ABB RAPID module: MAIN_1.mod

MODULE MAIN_1
GLOBAL VAR robtarget robpoint0 = p:{{1015.000, 0.000, 1372.000}, {0.707107, 0.000000, 0.707107, 0.000000}, 0}{cfg 0, 0, -1, 0, 0, -1, 0, 0}{Ej 0,0,0,0,0,0}
GLOBAL VAR robtarget robpoint1 = p:{{1015.000, 0.000, 1272.000}, {0.707107, 0.000000, 0.707107, 0.000000}, 0}{cfg 0, 0, -1, 0, -1, 0, 0, 1}{Ej 0,0,0,0,0,0}
GLOBAL VAR robtarget robpoint2 = p:{{187.264, 125.487, 305.356}, {0.001606, 0.000000, 0.999999, -0.000000}, 0}{cfg -1, 0, -1, 0, 0, -1, 0, 0}{Ej 0,0,0,0,0,0}
GLOBAL VAR robtarget robpoint3 = p:{{187.786, 125.499, 139.112}, {0.001571, -0.000026, 0.999999, 0.000035}, 0}{cfg -1, 0, -1, 0, 0, -1, 0, 0}{Ej 0,0,0,0,0,0}
GLOBAL VAR robtarget robpoint4 = p:{{187.272, 447.522, 305.347}, {0.001614, 0.000009, 0.999999, -0.000017}, 0}{cfg -1, 0, 0, 0, 0, -1, 0, 0}{Ej 0,0,0,0,0,0}
GLOBAL VAR robtarget robpoint5 = p:{{187.851, 447.517, 126.235}, {0.001614, 0.000009, 0.999999, -0.000017}, 0}{cfg -1, 0, 0, 0, 0, -1, 0, 0}{Ej 0,0,0,0,0,0}
GLOBAL VAR robtarget robpoint6 = p:{{187.272, 447.522, 305.347}, {0.001614, 0.000009, 0.999999, -0.000017}, 0}{cfg -1, 0, 0, 0, 0, -1, 0, 0}{Ej 0,0,0,0,0,0}
GLOBAL VAR robtarget robpoint7 = p:{{312.208, 292.214, 255.156}, {0.086206, -0.385314, 0.917581, 0.046341}, 0}{cfg 0, 0, 0, 0, 0, -2, 0, 0}{Ej 0,0,0,0,0,0}
GLOBAL VAR robtarget robpoint8 = p:{{430.047, 43.774, 231.503}, {0.086206, -0.385314, 0.917581, 0.046341}, 0}{cfg 0, 0, -1, 0, 0, -2, 0, 0}{Ej 0,0,0,0,0,0}
GLOBAL VAR robtarget robpoint9 = p:{{109.688, -153.222, 161.073}, {0.086206, -0.385314, 0.917581, 0.046341}, 0}{cfg 0, 0, 0, 0, 0, -2, 0, 0}{Ej 0,0,0,0,0,0}
GLOBAL VAR robtarget robpoint10 = p:{{312.208, 292.214, 255.156}, {0.086206, -0.385314, 0.917581, 0.046341}, 0}{cfg 0, 0, 0, 0, 0, -2, 0, 0}{Ej 0,0,0,0,0,0}
GLOBAL VAR robtarget robpoint11 = p:{{19.898, 201.357, 302.721}, {0.032125, 0.675431, -0.735891, 0.034999}, 0}{cfg 0, 0, -1, -1, 0, 0, 0, 0}{Ej 0,0,0,0,0,0}
GLOBAL VAR robtarget robpoint12 = p:{{19.898, 174.307, 19.008}, {0.032125, 0.675431, -0.735891, 0.034999}, 0}{cfg 0, 0, 0, -1, 0, 0, 0, 0}{Ej 0,0,0,0,0,0}
GLOBAL VAR robtarget robpoint13 = p:{{378.402, 174.416, 18.997}, {0.032125, 0.675431, -0.735891, 0.034999}, 0}{cfg 0, 0, -1, 0, 0, -1, 0, 0}{Ej 0,0,0,0,0,0}
GLOBAL VAR robtarget robpoint14 = p:{{380.996, 112.363, 34.882}, {0.106872, 0.666888, -0.728163, 0.116691}, 0}{cfg 0, 0, 0, -1, 0, -1, 0, 0}{Ej 0,0,0,0,0,0}
GLOBAL VAR robtarget robpoint15 = p:{{16.551, 114.359, 34.226}, {0.106872, 0.666888, -0.728163, 0.116691}, 0}{cfg 0, 0, 0, -1, 0, 0, 0, 0}{Ej 0,0,0,0,0,0}
GLOBAL VAR robtarget robpoint16 = p:{{26.434, 54.524, 46.072}, {0.025638, -0.672233, 0.739358, 0.028195}, 0}{cfg 0, 0, 0, -1, 0, 0, 0, 0}{Ej 0,0,0,0,0,0}
GLOBAL VAR robtarget robpoint17 = p:{{385.448, 48.050, 45.137}, {0.065816, -0.669242, 0.736571, 0.072433}, 0}{cfg 0, 0, 0, 0, 0, -1, 0, 0}{Ej 0,0,0,0,0,0}
GLOBAL VAR robtarget robpoint18 = p:{{385.448, -1.625, 295.251}, {0.065816, -0.669242, 0.736571, 0.072433}, 0}{cfg 0, 0, 0, 0, 0, -1, 0, 0}{Ej 0,0,0,0,0,0}
GLOBAL VAR robtarget robpoint19 = p:{{-49.939, 252.644, 419.997}, {0.002333, -0.707103, 0.707104, 0.002024}, 0}{cfg -1, 0, 0, 0, 0, -2, 0, 0}{Ej 0,0,0,0,0,0}
GLOBAL VAR robtarget robpoint20 = p:{{-49.895, 253.259, 319.999}, {0.002333, -0.707103, 0.707104, 0.002024}, 0}{cfg -1, 0, 0, 0, 0, -2, 0, 0}{Ej 0,0,0,0,0,0}
GLOBAL VAR robtarget robpoint21 = p:{{0.000, 250.000, 270.000}, {0.002333, -0.707103, 0.707104, 0.002024}, 0}{cfg -1, 0, 0, 0, 0, -2, 0, 0}{Ej 0,0,0,0,0,0}
GLOBAL VAR robtarget robpoint22 = p:{{35.579, 247.455, 270.000}, {0.002592, -0.707102, 0.707105, 0.001666}, 0}{cfg -1, 0, 0, 0, 0, -2, 0, 0}{Ej 0,0,0,0,0,0}
GLOBAL VAR robtarget robpoint23 = p:{{70.433, 239.873, 270.000}, {0.002808, -0.707107, 0.707099, 0.001277}, 0}{cfg -1, 0, 0, 0, 0, -2, 0, 0}{Ej 0,0,0,0,0,0}
GLOBAL VAR robtarget robpoint24 = p:{{103.854, 227.408, 270.000}, {0.002956, -0.707107, 0.707100, 0.000870}, 0}{cfg -1, 0, 0, 0, 0, -2, 0, 0}{Ej 0,0,0,0,0,0}
GLOBAL VAR robtarget robpoint25 = p:{{135.160, 210.313, 270.000}, {0.003054, -0.707106, 0.707100, 0.000438}, 0}{cfg -1, 0, 0, 0, 0, -2, 0, 0}{Ej 0,0,0,0,0,0}
GLOBAL VAR robtarget robpoint26 = p:{{163.715, 188.937, 270.000}, {0.003085, -0.707106, 0.707101, 0.000000}, 0}{cfg -1, 0, 0, 0, 0, -2, 0, 0}{Ej 0,0,0,0,0,0}
GLOBAL VAR robtarget robpoint27 = p:{{188.937, 163.715, 270.000}, {0.003054, -0.707106, 0.707100, -0.000438}, 0}{cfg -1, 0, 0, 0, 0, -2, 0, 0}{Ej 0,0,0,0,0,0}
GLOBAL VAR robtarget robpoint28 = p:{{210.313, 135.160, 270.000}, {0.002968, -0.707107, 0.707100, -0.000870}, 0}{cfg -1, 0, 0, 0, 0, -2, 0, 0}{Ej 0,0,0,0,0,0}
GLOBAL VAR robtarget robpoint29 = p:{{227.408, 103.854, 270.000}, {0.002814, -0.707107, 0.707099, -0.001284}, 0}{cfg -1, 0, 0, 0, 0, -2, 0, 0}{Ej 0,0,0,0,0,0}
GLOBAL VAR robtarget robpoint30 = p:{{239.873, 70.433, 270.000}, {0.002598, -0.707102, 0.707105, -0.001672}, 0}{cfg -1, 0, 0, 0, 0, -2, 0, 0}{Ej 0,0,0,0,0,0}
GLOBAL VAR robtarget robpoint31 = p:{{247.455, 35.579, 270.000}, {0.002333, -0.707103, 0.707104, -0.002024}, 0}{cfg -1, 0, 0, 0, 0, -2, 0, 0}{Ej 0,0,0,0,0,0}
GLOBAL VAR robtarget robpoint32 = p:{{250.000, 0.000, 270.000}, {0.002024, -0.707104, 0.707103, -0.002333}, 0}{cfg -1, 0, 0, 0, 0, -2, 0, 0}{Ej 0,0,0,0,0,0}
GLOBAL VAR robtarget robpoint33 = p:{{247.455, -35.579, 270.000}, {0.001672, -0.707105, 0.707102, -0.002598}, 0}{cfg -1, 0, 0, 0, 0, -2, 0, 0}{Ej 0,0,0,0,0,0}
GLOBAL VAR robtarget robpoint34 = p:{{239.873, -70.433, 270.000}, {0.001284, -0.707099, 0.707107, -0.002814}, 0}{cfg -2, 0, 0, 0, 0, -2, 0, 0}{Ej 0,0,0,0,0,0}
GLOBAL VAR robtarget robpoint35 = p:{{227.408, -103.854, 270.000}, {0.000870, -0.707100, 0.707107, -0.002968}, 0}{cfg -2, 0, 0, 0, 0, -2, 0, 0}{Ej 0,0,0,0,0,0}
GLOBAL VAR robtarget robpoint36 = p:{{210.313, -135.160, 270.000}, {0.000438, -0.707100, 0.707106, -0.003054}, 0}{cfg -2, 0, 0, 0, 0, -2, 0, 0}{Ej 0,0,0,0,0,0}
GLOBAL VAR robtarget robpoint37 = p:{{188.937, -163.715, 270.000}, {0.000000, -0.707101, 0.707106, -0.003085}, 0}{cfg -2, 0, 0, 0, 0, -2, 0, 0}{Ej 0,0,0,0,0,0}
GLOBAL VAR robtarget robpoint38 = p:{{163.715, -188.937, 270.000}, {0.000438, 0.707100, -0.707106, 0.003054}, 0}{cfg -2, 0, 0, 0, 0, -2, 0, 0}{Ej 0,0,0,0,0,0}
GLOBAL VAR robtarget robpoint39 = p:{{135.160, -210.313, 270.000}, {0.000870, 0.707100, -0.707107, 0.002968}, 0}{cfg -2, 0, 0, 0, 0, -2, 0, 0}{Ej 0,0,0,0,0,0}
GLOBAL VAR robtarget robpoint40 = p:{{103.854, -227.408, 270.000}, {0.001284, 0.707099, -0.707107, 0.002814}, 0}{cfg -2, 0, 0, 0, 0, -2, 0, 0}{Ej 0,0,0,0,0,0}
GLOBAL VAR robtarget robpoint41 = p:{{70.433, -239.873, 270.000}, {0.001672, 0.707105, -0.707102, 0.002598}, 0}{cfg -2, 0, 0, 0, 0, -2, 0, 0}{Ej 0,0,0,0,0,0}
GLOBAL VAR robtarget robpoint42 = p:{{35.579, -247.455, 270.000}, {0.002024, 0.707104, -0.707103, 0.002333}, 0}{cfg -2, 0, 0, 0, 0, -2, 0, 0}{Ej 0,0,0,0,0,0}
GLOBAL VAR robtarget robpoint43 = p:{{0.000, -250.000, 270.000}, {0.002024, 0.707104, -0.707103, 0.002333}, 0}{cfg -2, 0, 0, 0, 0, -2, 0, 0}{Ej 0,0,0,0,0,0}
GLOBAL VAR robtarget robpoint44 = p:{{0.000, -250.000, 270.000}, {0.002333, 0.707103, -0.707104, 0.002024}, 0}{cfg -2, 0, 0, 0, 0, -2, 0, 0}{Ej 0,0,0,0,0,0}
GLOBAL VAR robtarget robpoint45 = p:{{-35.579, -247.455, 270.000}, {0.002598, 0.707102, -0.707105, 0.001672}, 0}{cfg -2, 0, 0, 0, 0, -2, 0, 0}{Ej 0,0,0,0,0,0}
GLOBAL VAR robtarget robpoint46 = p:{{-70.433, -239.873, 270.000}, {0.002808, 0.707107, -0.707099, 0.001277}, 0}{cfg -2, 0, 0, 0, 0, -2, 0, 0}{Ej 0,0,0,0,0,0}
GLOBAL VAR robtarget robpoint47 = p:{{-103.854, -227.408, 270.000}, {0.002956, 0.707107, -0.707100, 0.000870}, 0}{cfg -2, 0, 0, 0, 0, -2, 0, 0}{Ej 0,0,0,0,0,0}
GLOBAL VAR robtarget robpoint48 = p:{{-135.160, -210.313, 270.000}, {0.003054, 0.707106, -0.707100, 0.000438}, 0}{cfg -2, 0, 0, 0, 0, -2, 0, 0}{Ej 0,0,0,0,0,0}
GLOBAL VAR robtarget robpoint49 = p:{{-163.715, -188.937, 270.000}, {0.003085, 0.707106, -0.707101, 0.000000}, 0}{cfg -2, 0, 0, 0, 0, -2, 0, 0}{Ej 0,0,0,0,0,0}
GLOBAL VAR robtarget robpoint50 = p:{{-188.937, -163.715, 270.000}, {0.003054, 0.707106, -0.707100, -0.000438}, 0}{cfg -2, 0, 0, 0, 0, -2, 0, 0}{Ej 0,0,0,0,0,0}
GLOBAL VAR robtarget robpoint51 = p:{{-210.313, -135.160, 270.000}, {0.002956, 0.707107, -0.707100, -0.000870}, 0}{cfg -2, 0, 0, 0, 0, -2, 0, 0}{Ej 0,0,0,0,0,0}
GLOBAL VAR robtarget robpoint52 = p:{{-227.408, -103.854, 270.000}, {0.002801, 0.707107, -0.707099, -0.001284}, 0}{cfg -2, 0, 0, 0, 0, -2, 0, 0}{Ej 0,0,0,0,0,0}
GLOBAL VAR robtarget robpoint53 = p:{{-239.873, -70.433, 270.000}, {0.002598, 0.707102, -0.707105, -0.001672}, 0}{cfg -2, 0, 0, 0, 0, -2, 0, 0}{Ej 0,0,0,0,0,0}
GLOBAL VAR robtarget robpoint54 = p:{{-247.455, -35.579, 270.000}, {0.002333, 0.707103, -0.707104, -0.002024}, 0}{cfg -1, 0, 0, 0, 0, -2, 0, 0}{Ej 0,0,0,0,0,0}
GLOBAL VAR robtarget robpoint55 = p:{{-250.000, 0.000, 270.000}, {0.002024, 0.707104, -0.707103, -0.002333}, 0}{cfg -1, 0, 0, 0, 0, -2, 0, 0}{Ej 0,0,0,0,0,0}
GLOBAL VAR robtarget robpoint56 = p:{{-247.455, 35.579, 270.000}, {0.001666, 0.707105, -0.707102, -0.002592}, 0}{cfg -1, 0, 0, 0, 0, -2, 0, 0}{Ej 0,0,0,0,0,0}
GLOBAL VAR robtarget robpoint57 = p:{{-239.873, 70.433, 270.000}, {0.001284, 0.707099, -0.707107, -0.002801}, 0}{cfg -1, 0, 0, 0, 0, -2, 0, 0}{Ej 0,0,0,0,0,0}
GLOBAL VAR robtarget robpoint58 = p:{{-227.408, 103.854, 270.000}, {0.000870, 0.707100, -0.707107, -0.002968}, 0}{cfg -1, 0, 0, 0, 0, -2, 0, 0}{Ej 0,0,0,0,0,0}
GLOBAL VAR robtarget robpoint59 = p:{{-210.313, 135.160, 270.000}, {0.000438, 0.707100, -0.707106, -0.003054}, 0}{cfg -1, 0, 0, 0, 0, -2, 0, 0}{Ej 0,0,0,0,0,0}
GLOBAL VAR robtarget robpoint60 = p:{{-188.937, 163.715, 270.000}, {0.000000, -0.707101, 0.707106, 0.003085}, 0}{cfg -1, 0, 0, 0, 0, -2, 0, 0}{Ej 0,0,0,0,0,0}
GLOBAL VAR robtarget robpoint61 = p:{{-163.715, 188.937, 270.000}, {0.000438, -0.707100, 0.707106, 0.003054}, 0}{cfg -1, 0, 0, 0, 0, -2, 0, 0}{Ej 0,0,0,0,0,0}
GLOBAL VAR robtarget robpoint62 = p:{{-135.160, 210.313, 270.000}, {0.000870, -0.707100, 0.707107, 0.002956}, 0}{cfg -1, 0, 0, 0, 0, -2, 0, 0}{Ej 0,0,0,0,0,0}
GLOBAL VAR robtarget robpoint63 = p:{{-103.854, 227.408, 270.000}, {0.001284, -0.707099, 0.707107, 0.002814}, 0}{cfg -1, 0, 0, 0, 0, -2, 0, 0}{Ej 0,0,0,0,0,0}
GLOBAL VAR robtarget robpoint64 = p:{{-70.433, 239.873, 270.000}, {0.001672, -0.707105, 0.707102, 0.002598}, 0}{cfg -1, 0, 0, 0, 0, -2, 0, 0}{Ej 0,0,0,0,0,0}
GLOBAL VAR robtarget robpoint65 = p:{{-35.579, 247.455, 270.000}, {0.002024, -0.707104, 0.707103, 0.002333}, 0}{cfg -1, 0, 0, 0, 0, -2, 0, 0}{Ej 0,0,0,0,0,0}
GLOBAL VAR robtarget robpoint66 = p:{{0.000, 250.000, 270.000}, {0.002024, -0.707104, 0.707103, 0.002333}, 0}{cfg -1, 0, 0, 0, 0, -2, 0, 0}{Ej 0,0,0,0,0,0}
GLOBAL VAR robtarget robpoint67 = p:{{49.895, 253.258, 319.999}, {0.002024, -0.707104, 0.707103, 0.002333}, 0}{cfg -1, 0, 0, 0, 0, -2, 0, 0}{Ej 0,0,0,0,0,0}
GLOBAL VAR robtarget robpoint68 = p:{{49.939, 252.642, 419.997}, {0.002024, -0.707104, 0.707103, 0.002333}, 0}{cfg -1, 0, 0, 0, 0, -2, 0, 0}{Ej 0,0,0,0,0,0}
GLOBAL VAR robtarget robpoint69 = p:{{187.264, 125.487, 305.356}, {0.001606, 0.000000, 0.999999, -0.000000}, 0}{cfg -1, 0, -1, 0, 0, -1, 0, 0}{Ej 0,0,0,0,0,0}
GLOBAL VAR robtarget robpoint70 = p:{{187.786, 125.499, 139.112}, {0.001571, -0.000026, 0.999999, 0.000035}, 0}{cfg -1, 0, -1, 0, 0, -1, 0, 0}{Ej 0,0,0,0,0,0}
GLOBAL VAR robtarget robpoint71 = p:{{187.264, 125.487, 305.356}, {0.001606, 0.000000, 0.999999, -0.000000}, 0}{cfg -1, 0, -1, 0, 0, -1, 0, 0}{Ej 0,0,0,0,0,0}

GLOBAL VAR robtarget robpoint72 = p:{{1015.000, -1000.000, 1237.000}, {0.707107, 0.000000, 0.707107, -0.000000}, 0}{cfg -1, 0, 0, 0, 0, -1, 0, 0}{Ej 0,0,0,0,0,0}

GLOBAL Proc main()
    MoveJ robpoint0,v50,z50,tool03,wobj16
    MoveL robpoint1,v50,z50,tool03,wobj16
    SetDO D_OUT_5, 1;
    SetDO D_OUT_5, 1;
    SetDO D_OUT_5, 0.5;
    SetDO D_OUT_5, true;
    SetDO D_OUT_5, 1;
    SetDO D_OUT_5, 1;
    SetDO D_OUT_5, 0.5;
    SetDO D_OUT_5, true;
    SetDO var, val;
    SetDO var, val;
    WaitDI D_IN_5, 1;
    WaitDI D_IN_5, 1;
    WaitDI D_IN_5, 0.5;
    WaitDI D_IN_5, true;
    WaitDI D_IN_5, 1, \MaxTime:=0.1;
    WaitDI var, val;
    WaitDI var, val, \MaxTime:=0.1;
    TPWrite "Message";
    REMOTE_PROG_CALL_171;
    CODE_INSERT_172
    wobj16.x = 719.013
    wobj16.y = -664.003
    wobj16.z = 0.000
    wobj16.q1 = 1.000000
    wobj16.q2 = 0.000000
    wobj16.q3 = 0.000000
    wobj16.q4 = 0.000000
    tool03.x = 129.073
    tool03.y = 0.000
    tool03.z = 85.477
    tool03.q1 = 0.980187
    tool03.q2 = 0.000000
    tool03.q3 = 0.198076
    tool03.q4 = 0.000000
    MoveJ robpoint2,v50,z10,tool03,wobj16
    MoveL robpoint3,v100,fine,tool03,wobj16
    SetDO D_OUT_5, 1;
    PICK_PART_111;
    MoveL robpoint4,v300,z10,tool03,wobj16
    MoveL robpoint5,v100,fine,tool03,wobj16
    SetDO D_OUT_5, 0;
    PLACE_PART_112;
    MoveL robpoint6,v100,z10,tool03,wobj16
    wobj16.x = 577.67
    wobj16.y = 392.250
    wobj16.z = 0.000
    wobj16.q1 = 0.942759
    wobj16.q2 = 0.000000
    wobj16.q3 = 0.000000
    wobj16.q4 = 0.333474
    MoveJ robpoint7,v100,z25,tool03,wobj16
    MoveC robpoint8,robpoint9,v100,z25,tool03,wobj16
    MoveL robpoint10,v100,fine,tool03,wobj16
    wobj16.x = 0
    wobj16.y = 782.714
    wobj16.z = 377.610
    wobj16.q1 = 1.000000
    wobj16.q2 = 0.000000
    wobj16.q3 = 0.000000
    wobj16.q4 = 0.000000
    MoveJ robpoint11,v100,fine,tool03,wobj16
    MoveL robpoint12,v100,fine,tool03,wobj16
    MoveL robpoint13,v100,fine,tool03,wobj16
    MoveL robpoint14,v100,fine,tool03,wobj16
    MoveL robpoint15,v100,fine,tool03,wobj16
    MoveL robpoint16,v100,fine,tool03,wobj16
    MoveL robpoint17,v100,fine,tool03,wobj16
    MoveL robpoint18,v100,fine,tool03,wobj16
    EVENT_PROG_START_101;
    wobj16.x = 13.637
    wobj16.y = -840.080
    wobj16.z = 0.000
    wobj16.q1 = 0.707107
    wobj16.q2 = 0.000000
    wobj16.q3 = 0.000000
    wobj16.q4 = -0.707107
    MoveJ robpoint19,v1000,z1,tool03,wobj16
    EVENT_PATH_APPROACH_102;
    MoveL robpoint20,v1000,z1,tool03,wobj16
    MoveL robpoint21,v1000,z1,tool03,wobj16
    EVENT_PATH_START_103;
    MoveL robpoint22,v50,z1,tool03,wobj16
    MoveL robpoint23,v50,z1,tool03,wobj16
    MoveL robpoint24,v50,z1,tool03,wobj16
    MoveL robpoint25,v50,z1,tool03,wobj16
    MoveL robpoint26,v50,z1,tool03,wobj16
    MoveL robpoint27,v50,z1,tool03,wobj16
    MoveL robpoint28,v50,z1,tool03,wobj16
    MoveL robpoint29,v50,z1,tool03,wobj16
    MoveL robpoint30,v50,z1,tool03,wobj16
    MoveL robpoint31,v50,z1,tool03,wobj16
    MoveL robpoint32,v50,z1,tool03,wobj16
    MoveL robpoint33,v50,z1,tool03,wobj16
    MoveL robpoint34,v50,z1,tool03,wobj16
    MoveL robpoint35,v50,z1,tool03,wobj16
    MoveL robpoint36,v50,z1,tool03,wobj16
    MoveL robpoint37,v50,z1,tool03,wobj16
    MoveL robpoint38,v50,z1,tool03,wobj16
    MoveL robpoint39,v50,z1,tool03,wobj16
    MoveL robpoint40,v50,z1,tool03,wobj16
    MoveL robpoint41,v50,z1,tool03,wobj16
    MoveL robpoint42,v50,z1,tool03,wobj16
    MoveL robpoint43,v50,z1,tool03,wobj16
    MoveL robpoint44,v50,z1,tool03,wobj16
    MoveL robpoint45,v50,z1,tool03,wobj16
    MoveL robpoint46,v50,z1,tool03,wobj16
    MoveL robpoint47,v50,z1,tool03,wobj16
    MoveL robpoint48,v50,z1,tool03,wobj16
    MoveL robpoint49,v50,z1,tool03,wobj16
    MoveL robpoint50,v50,z1,tool03,wobj16
    MoveL robpoint51,v50,z1,tool03,wobj16
    MoveL robpoint52,v50,z1,tool03,wobj16
    MoveL robpoint53,v50,z1,tool03,wobj16
    MoveL robpoint54,v50,z1,tool03,wobj16
    MoveL robpoint55,v50,z1,tool03,wobj16
    MoveL robpoint56,v50,z1,tool03,wobj16
    MoveL robpoint57,v50,z1,tool03,wobj16
    MoveL robpoint58,v50,z1,tool03,wobj16
    MoveL robpoint59,v50,z1,tool03,wobj16
    MoveL robpoint60,v50,z1,tool03,wobj16
    MoveL robpoint61,v50,z1,tool03,wobj16
    MoveL robpoint62,v50,z1,tool03,wobj16
    MoveL robpoint63,v50,z1,tool03,wobj16
    MoveL robpoint64,v50,z1,tool03,wobj16
    MoveL robpoint65,v50,z1,tool03,wobj16
    MoveL robpoint66,v50,z1,tool03,wobj16
    EVENT_PATH_FINISH_105;
    MoveL robpoint67,v1000,z1,tool03,wobj16
    MoveL robpoint68,v1000,z1,tool03,wobj16
    EVENT_PATH_RETRACT_106;
    EVENT_PROG_FINISH_107;
    wobj16.x = 719.013
    wobj16.y = -664.003
    wobj16.z = 0.000
    wobj16.q1 = 1.000000
    wobj16.q2 = 0.000000
    wobj16.q3 = 0.000000
    wobj16.q4 = 0.000000
    MoveJ robpoint69,v1000,z1,tool03,wobj16
    Wait 1.250
    MoveL robpoint70,v1000,z1,tool03,wobj16
    WaitDI D_IN_1, 1;
    MoveL robpoint71,v1000,z1,tool03,wobj16
    PROG1_withaverylongnameandspecialcharacters;
EndProc
EndModule
GLOBAL Proc main()
    wobj16.x = 0
    wobj16.y = 1000.000
    wobj16.z = 0.000
    wobj16.q1 = 1.000000
    wobj16.q2 = 0.000000
    wobj16.q3 = 0.000000
    wobj16.q4 = 0.000000
    tool03.x = 0.000
    tool03.y = 0.000
    tool03.z = 200.000
    tool03.q1 = 1.000000
    tool03.q2 = 0.000000
    tool03.q3 = 0.000000
    tool03.q4 = 0.000000
    MoveJ robpoint72,v1000,z1,tool03,wobj16
EndProc
EndModule
